Fanuc KAREL source: KD00040.KL

PROGRAM KD00040
%NOLOCKGROUP
VAR
  I: INTEGER
  J: INTEGER
  B: BOOLEAN
  R: REAL
  S: STRING[80]
  PTH: PATH
BEGIN
  WRITE(PTH)
END KD00040
